Fanuc KAREL source: KC00018.KL

PROGRAM KC00018
%NOLOCKGROUP
%ENVIRONMENT BYNAM
VAR
  I: INTEGER
  J: INTEGER
  K: INTEGER
  R: REAL
  B: BOOLEAN
  S: STRING[80]
  T: STRING[80]
  P: PATH
  Q: PATH
  AI: ARRAY[8] OF INTEGER
  AB: ARRAY[244] OF BYTE
BEGIN
  VAR_INFO(S,T,B,S,I,AI,J,K)
END KC00018
